FUNCTION_BLOCK EV_Template (* TEMPLATE for the report form of your equipment, EV_<Equipment>: copy it under that name, then change what says YOUR OWN, and this comment; keep the rest as it is. Names the equipment's two channels, and unpacks its state channel into named values (its inputs and who holds it) for a skill. Technical: Names Template's channels; typed view of its state channel (inputs and holder) *)
  (* Standard: 61499-2 *)
  (* Version 0.1, 2026-09-28, Project contributors, AAU Smart Production Lab *)
  PACKAGE capping;
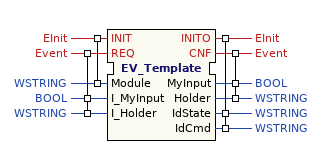
  EVENT_INPUT
    INIT : EInit WITH Module; (* Name the equipment's channels *)
    REQ WITH I_MyInput, I_Holder; (* The equipment's state arrived *)
  END_EVENT
  EVENT_OUTPUT
    INITO : EInit WITH IdState, IdCmd; (* IdState and IdCmd are set *)
    CNF WITH MyInput, Holder; (* The values below are updated *)
  END_EVENT
  VAR_INPUT
    Module : WSTRING; (* The module's name; its local channels are named after it (loc[<Module>/...]) *)
    I_MyInput : BOOL; (* YOUR OWN, one per input pin. MyInput as read or received *)
    I_Holder : WSTRING; (* Holder as read or received *)
  END_VAR
  VAR_OUTPUT
    MyInput : BOOL; (* YOUR OWN, one per input pin. Template: MyInput, an input *)
    Holder : WSTRING; (* Who holds the equipment (empty: free) *)
    IdState : WSTRING; (* Local channel of the equipment's state *)
    IdCmd : WSTRING; (* Local channel of the equipment's commands *)
  END_VAR
  EC_STATES
    INIT : INIT -> INITO;
    REQ : REQ -> CNF;
  END_STATES
  ALGORITHM INIT IN ST:
IdState := CONCAT(CONCAT("loc[", Module), "/Template/state]");  (* YOUR OWN: the equipment item's name, as Name in EQ_ *)
IdCmd := CONCAT(CONCAT("loc[", Module), "/Template/cmd]");  (* YOUR OWN: the equipment item's name, as Name in EQ_ *)
  END_ALGORITHM
  ALGORITHM REQ IN ST:
MyInput := I_MyInput;  (* YOUR OWN: one line per input pin *)
Holder := I_Holder;
  END_ALGORITHM
END_FUNCTION_BLOCK
